(* IEC 61131-3 sources: plc-cip-batch-control/plc/types, 3 files *)

(* ---- Types_Cip.st ---- *)
(*
    Types_Cip.st: data types for the CIP skid controller.

    Naming follows the usual IEC prefixes: x BOOL, i INT, r REAL, t TIME,
    s STRING, e enumeration, st structure, fb function block instance.

    Enumeration members are prefixed because IEC 61131-3 puts them in the
    global namespace and PH_IDLE and UST_IDLE are different things.
*)

TYPE
    (* ISA-88 procedural state model, trimmed to the states this unit uses. *)
    E_UnitState : (
        UST_IDLE        := 0,
        UST_STARTING    := 1,
        UST_RUNNING     := 2,
        UST_HOLDING     := 3,
        UST_HELD        := 4,
        UST_RESTARTING  := 5,
        UST_COMPLETING  := 6,
        UST_COMPLETE    := 7,
        UST_ABORTING    := 8,
        UST_ABORTED     := 9
    );

    (* The CIP procedure. Phases run in this order; the recipe may skip some. *)
    E_Phase : (
        PH_IDLE                := 0,
        PH_PRE_RINSE           := 1,
        PH_CAUSTIC_WASH        := 2,
        PH_INTERMEDIATE_RINSE  := 3,
        PH_ACID_WASH           := 4,
        PH_FINAL_RINSE         := 5,
        PH_SANITISE            := 6,
        PH_COMPLETE            := 7
    );

    (* Every phase runs the same four steps; only its parameters differ. *)
    E_PhaseStep : (
        PS_IDLE      := 0,
        PS_LINEUP    := 1,
        PS_CHARGE    := 2,
        PS_CIRCULATE := 3,
        PS_RECOVER   := 4,
        PS_DONE      := 5
    );

    E_Source : (
        SRC_NONE       := 0,
        SRC_FRESH      := 1,
        SRC_RECOVERED  := 2,
        SRC_CAUSTIC    := 3,
        SRC_ACID       := 4
    );

    E_Return : (
        RET_DRAIN     := 0,
        RET_RECOVERY  := 1,
        RET_CAUSTIC   := 2,
        RET_ACID      := 3,
        RET_BALANCE   := 4
    );

    E_FailCode : (
        FC_NONE             := 0,
        FC_LINEUP_TIMEOUT   := 1,
        FC_CHARGE_TIMEOUT   := 2,
        FC_TEMP_TIMEOUT     := 3,
        FC_PHASE_TIMEOUT    := 4,
        FC_FLOW_LOW         := 5,
        FC_PUMP_FAULT       := 6,
        FC_OPERATOR_ABORT   := 7,
        FC_SAFETY_TRIP      := 8,
        FC_RINSE_NOT_CLEAN  := 9,
        FC_LEVEL_LOW        := 10,
        FC_SENSOR_FAULT     := 11
    );
END_TYPE

TYPE
    (*
        What one phase has to achieve. PRG_Sequence fills this from the recipe
        and hands it to the single phase engine, so adding a phase is a matter
        of parameters rather than another copy of the same logic.
    *)
    ST_PhaseParams : STRUCT
        eSource         : E_Source;
        eReturn         : E_Return;
        rTempSp         : REAL;     (* heat setpoint, degC *)
        rTempMin        : REAL;     (* below this the hold timer does not count *)
        rConcSp         : REAL;     (* chemical strength, % w/w *)
        rConcMin        : REAL;
        rConcMax        : REAL;
        rFlowSp         : REAL;     (* m3/h *)
        rFlowMin        : REAL;     (* below this the hold timer does not count *)
        tHold           : TIME;     (* verified hold required to pass *)
        tMinPhase       : TIME;
        tMaxPhase       : TIME;
        tRecover        : TIME;     (* push the circuit contents back or to drain *)
        xHeat           : BOOL;
        xDose           : BOOL;
        xRecirculate    : BOOL;     (* closed loop through the balance tank *)
        xAdaptiveEnd    : BOOL;     (* terminate on the return conductivity *)
        rEndConductivity : REAL;    (* mS/cm, adaptive rinses only *)
    END_STRUCT

    (* What the phase engine asks the control layer to do this scan. *)
    ST_Demand : STRUCT
        eSource      : E_Source;
        eReturn      : E_Return;
        rFlowSp      : REAL;
        rTempSp      : REAL;
        xHeat        : BOOL;
        xDose        : BOOL;
        xSupplyPump  : BOOL;
        xReturnPump  : BOOL;
        xFillValve   : BOOL;
    END_STRUCT

    (* One line of the electronic batch record. *)
    ST_PhaseResult : STRUCT
        ePhase           : E_Phase;
        xExecuted        : BOOL;
        xPass            : BOOL;
        eFail            : E_FailCode;
        rDurationS       : REAL;
        rHoldAchievedS   : REAL;
        rHoldRequiredS   : REAL;    (* zero when the endpoint is the conductivity *)
        xAdaptiveEnd     : BOOL;
        rMinTempC        : REAL := 999.0;
        rMaxTempC        : REAL;
        rMeanConcPct     : REAL;
        rMinFlow         : REAL := 999.0;
        rWaterL          : REAL;
        rChemL           : REAL;
        rEnergyKWh       : REAL;
        rEndConductivity : REAL;
    END_STRUCT

    ST_Recipe : STRUCT
        sName            : STRING[24] := 'default';
        xUseAcid         : BOOL := TRUE;
        xUseSanitise     : BOOL := FALSE;
        xAdaptive        : BOOL := FALSE;
        rFlowSp          : REAL := 18.0;
        tPreRinse        : TIME := T#3m;
        rCausticTempSp   : REAL := 75.0;
        rCausticTempMin  : REAL := 70.0;
        rCausticConcSp   : REAL := 2.0;
        tCausticHold     : TIME := T#10m;
        tIntRinse        : TIME := T#2m;
        rAcidTempSp      : REAL := 60.0;
        rAcidTempMin     : REAL := 55.0;
        rAcidConcSp      : REAL := 1.0;
        tAcidHold        : TIME := T#5m;
        tFinalRinse      : TIME := T#3m;
        rSanitiseTempSp  : REAL := 85.0;
        rSanitiseTempMin : REAL := 80.0;
        tSanitiseHold    : TIME := T#10m;
        rRinseEndCond    : REAL := 0.10;
        tPhaseMax        : TIME := T#45m;
        tRinseMax        : TIME := T#12m;   (* adaptive rinses fail rather than run on *)
        tRinseMin        : TIME := T#60s;   (* floor under the transport-delay blanking *)
        rFlowMin         : REAL := 14.0;
    END_STRUCT

    ST_Kpi : STRUCT
        rFreshWaterL     : REAL;
        rRecoveredWaterL : REAL;
        rEffluentL       : REAL;
        rCausticL        : REAL;
        rAcidL           : REAL;
        rEnergyKWh       : REAL;
        rCycleTimeS      : REAL;
        xVerifiedClean   : BOOL;
    END_STRUCT

    ST_Alarm : STRUCT
        xActive   : BOOL;
        xLatched  : BOOL;
        xAcked    : BOOL;
        iPriority : INT;
        rTimeInS  : REAL;
        iCount    : INT;
    END_STRUCT
END_TYPE

(* ---- GVL_Cip.st ---- *)
(*
    GVL_Cip.st: internal state shared between the five programs.

    Nothing here is located: these are the controller's own working data, not
    field I/O. PRG_Sequence owns the state and phase variables, PRG_Control owns
    the outputs, PRG_Alarms owns the alarm array and PRG_Kpi owns the totals.
    Every other program reads them.
*)

VAR_GLOBAL CONSTANT
    C_ALARM_COUNT       : INT  := 13;
    C_PHASE_COUNT       : INT  := 6;

    (* Alarm identifiers, used as the index into gAlarms. *)
    C_ALM_SAFETY        : INT  := 1;
    C_ALM_SUPPLY_PUMP   : INT  := 2;
    C_ALM_RETURN_PUMP   : INT  := 3;
    C_ALM_LEVEL_LOW     : INT  := 4;
    C_ALM_CAUSTIC_LOW   : INT  := 5;
    C_ALM_ACID_LOW      : INT  := 6;
    C_ALM_TEMP_LOW      : INT  := 7;
    C_ALM_FLOW_LOW      : INT  := 8;
    C_ALM_CIRCUIT_BUSY  : INT  := 9;
    C_ALM_PHASE_TIMEOUT : INT  := 10;
    C_ALM_NOT_CLEAN     : INT  := 11;
    C_ALM_NO_STEAM      : INT  := 12;
    C_ALM_COND_SENSOR   : INT  := 13;

    (* Skid geometry. The plant model holds the same figures; docs/model.md
       explains why they are stated twice and how the test keeps them equal. *)
    C_BALANCE_TANK_L    : REAL := 1200.0;
    C_CIRCUIT_VOLUME_L  : REAL := 450.0;    (* holdup of the circuit being cleaned *)
    (* A rinse endpoint cannot be believed until the return sensor has seen
       what was in the circuit when the rinse started. One and a half circuit
       turnovers is the blanking time. *)
    C_RINSE_TURNOVERS   : REAL := 1.5;
    C_FILL_TARGET_PCT   : REAL := 60.0;     (* recirculating phases *)
    (* Single-pass phases run the tank as a break volume at the lowest level
       the suction will stand. The rinse has to wash the tank out as well as
       the circuit and the tank washes out with a time constant of
       volume/flow: 156 litres at 18 m3/h is half a minute, 360 litres is
       nearly two and that difference is most of the rinse. *)
    C_RINSE_LEVEL_PCT   : REAL := 13.0;
    C_PUMP_START_PCT    : REAL := 10.0;     (* suction head to start the pump *)
    C_LEVEL_TRIP_PCT    : REAL := 7.0;
    C_CHEM_LEVEL_MIN    : REAL := 15.0;

    (* Two-point conductivity calibrations, mS/cm per % w/w, compensated to
       25 degC by the transmitter. Caustic is calibrated at 2 %, acid at 1 %. *)
    C_COND_K_CAUSTIC    : REAL := 47.0;
    C_COND_K_ACID       : REAL := 45.0;

    (* Positive-displacement dosing pumps, so the delivered volume is the
       valve-open time multiplied by a constant. *)
    C_CAUSTIC_DOSE_LPM  : REAL := 30.0;
    C_ACID_DOSE_LPM     : REAL := 20.0;

    C_TEMP_TOL          : REAL := 1.0;
    (* Plate-pack outlet limit. Above this the gaskets suffer and dissolved
       soil starts to bake onto the plates. *)
    C_SUPPLY_TEMP_LIMIT : REAL := 90.0;
    (* Task period. The harness asserts that the scan it runs matches. *)
    C_CYCLE_S           : REAL := 0.2;

    C_PUMP_SPEED_MIN    : REAL := 25.0;
    C_PUMP_SPEED_MAX    : REAL := 100.0;
END_VAR

VAR_GLOBAL
    (* ---- recipe and procedure state --------------------------------- *)
    gRecipe         : ST_Recipe;
    gUnitState      : E_UnitState;
    gPhase          : E_Phase;
    gPhaseStep      : E_PhaseStep;
    gFailCode       : E_FailCode;
    gPhaseParams    : ST_PhaseParams;
    gDemand         : ST_Demand;
    gResults        : ARRAY[1..6] OF ST_PhaseResult;
    gKpi            : ST_Kpi;
    giBatchId       : INT;

    (* ---- requests between programs ---------------------------------- *)
    gxSafetyTrip    : BOOL;     (* PRG_Safety -> everyone *)
    gxPermitRun     : BOOL;     (* PRG_Safety: it is safe to circulate *)
    gxPermitHeat    : BOOL;     (* PRG_Safety: steam may be admitted *)
    gxPermitDose    : BOOL;     (* PRG_Safety: chemical may be dosed *)
    gxHoldRequest   : BOOL;
    gxAbortRequest  : BOOL;
    gxPhaseExecute  : BOOL;
    gxPhaseDone     : BOOL;
    gxPhaseFailed   : BOOL;
    gxCycleReset    : BOOL;     (* one scan at the start of a batch *)
    gxPhaseStartPulse : BOOL;
    gxPhaseEndPulse : BOOL;
    giPhaseIndex    : INT;      (* which gResults entry the pulse refers to *)

    (* ---- derived measurements --------------------------------------- *)
    grConcentrationPct : REAL;  (* from the return conductivity *)
    grDeltaConductivity : REAL; (* return minus supply, the rinse criterion *)
    grCycleElapsedS : REAL;
    grPhaseElapsedS : REAL;
    grHoldAchievedS : REAL;
    grPlcTimeS      : REAL;     (* controller uptime, used to stamp alarms *)
    grCondFloor     : REAL;     (* reading the return must exceed in a wash *)
    gxCondSensorFault : BOOL;   (* the return element is not reading the process *)
    gxCondProven    : BOOL;     (* it saw the wash during this phase *)

    (* ---- alarms ------------------------------------------------------ *)
    gAlarms         : ARRAY[1..13] OF ST_Alarm;
    giFirstOut      : INT;
    giActiveAlarms  : INT;
    gxAlarmP1Active : BOOL;
END_VAR

(* ---- GVL_Io.st ---- *)
(*
    GVL_Io.st: the I/O image.

    These declarations are the single source of truth for the address map. The
    simulated field bus and the Modbus TCP server both build their tables by
    reading the AT addresses back out of the compiled program, so a tag cannot
    drift away from the address the logic uses. See docs/io_map.md.

    Address convention: %IXb.i is byte b bit i; %ID/%QD/%MD n is double word n.

    Inputs and outputs never share a number: inputs own bytes 0 and 1 and
    double words 0 to 15, outputs start at byte 2 and double word 16. IEC
    61131-3 keeps %I and %Q apart but some runtimes back both with one
    process image keyed by the number alone (RuSTy does, see
    docs/compiled_crosscheck.md); there %IX0.0 and %QX0.0 would be the same
    bit. Keeping the numbers disjoint costs nothing and works on both kinds.
*)

VAR_GLOBAL
    (* ---- digital inputs: plant status ------------------------------- *)
    xSafetyOk               AT %IX0.0 : BOOL;   (* safety relay healthy, E-stop clear *)
    xSupplyPumpRunning      AT %IX0.1 : BOOL;
    xReturnPumpRunning      AT %IX0.2 : BOOL;
    xSupplyPumpFault        AT %IX0.3 : BOOL;
    xReturnPumpFault        AT %IX0.4 : BOOL;
    xCircuitAvailable       AT %IX0.5 : BOOL;   (* the vessel is released for cleaning *)
    xSteamAvailable         AT %IX0.6 : BOOL;
    xBalanceTankLowLow      AT %IX0.7 : BOOL;   (* hard-wired float switch *)

    (* ---- operator commands -------------------------------------------
       These live in the memory area, not the input image, because they arrive
       from a panel or a SCADA client over the network rather than from a
       hard-wired button. The controller clears each one once it has taken the
       edge, so a client that writes a coil and forgets it still gets a pulse. *)
    xCmdStart               AT %MX0.0 : BOOL;
    xCmdHold                AT %MX0.1 : BOOL;
    xCmdRestart             AT %MX0.2 : BOOL;
    xCmdAbort               AT %MX0.3 : BOOL;
    xCmdReset               AT %MX0.4 : BOOL;
    xCmdAckAlarms           AT %MX0.5 : BOOL;

    (* ---- analogue inputs -------------------------------------------- *)
    rLevelBalanceTankPct    AT %ID0  : REAL;
    rTempSupplyC            AT %ID1  : REAL;    (* after the heat exchanger *)
    rTempReturnC            AT %ID2  : REAL;    (* back from the circuit *)
    rFlowSupplyM3h          AT %ID3  : REAL;
    rConductivityReturn     AT %ID4  : REAL;    (* mS/cm, temperature compensated *)
    rPressureSupplyBar      AT %ID5  : REAL;
    rLevelCausticPct        AT %ID6  : REAL;
    rLevelAcidPct           AT %ID7  : REAL;
    rLevelRecoveryPct       AT %ID8  : REAL;
    rConductivitySupply     AT %ID9  : REAL;    (* mS/cm, feed side *)
    rFlowMakeupM3h          AT %ID10 : REAL;    (* make-up into the balance tank *)
    rTempBalanceTankC       AT %ID11 : REAL;
    rConductivityTank       AT %ID12 : REAL;    (* CT-03, in the balance tank *)

    (* ---- digital outputs: valve matrix ------------------------------ *)
    xV01FreshWater          AT %QX2.0 : BOOL;
    xV02RecoveredWater      AT %QX2.1 : BOOL;
    xV03CausticDose         AT %QX2.2 : BOOL;
    xV04AcidDose            AT %QX2.3 : BOOL;
    xV05SupplyToCircuit     AT %QX2.4 : BOOL;
    xV06ReturnToDrain       AT %QX2.5 : BOOL;
    xV07ReturnToBalance     AT %QX2.6 : BOOL;
    xV08ReturnToCaustic     AT %QX2.7 : BOOL;
    xV09ReturnToRecovery    AT %QX3.0 : BOOL;
    xV10ReturnToAcid        AT %QX3.1 : BOOL;
    xSupplyPumpRun          AT %QX3.2 : BOOL;
    xReturnPumpRun          AT %QX3.3 : BOOL;
    xSteamIsolation         AT %QX3.4 : BOOL;
    xV11CausticSupply       AT %QX3.5 : BOOL;   (* caustic tank -> balance tank *)
    xV12AcidSupply          AT %QX3.6 : BOOL;

    (* ---- analogue outputs ------------------------------------------- *)
    rSupplyPumpSpeedPct     AT %QD16 : REAL;
    rSteamValvePct          AT %QD17 : REAL;

    (* ---- memory image published to SCADA ---------------------------- *)
    iHmiUnitState           AT %MW0 : INT;
    iHmiPhase               AT %MW1 : INT;
    iHmiPhaseStep           AT %MW2 : INT;
    iHmiFailCode            AT %MW3 : INT;
    iHmiActiveAlarms        AT %MW4 : INT;
    iHmiFirstOutAlarm       AT %MW5 : INT;
    iHmiBatchId             AT %MW6 : INT;

    rHmiFreshWaterL         AT %MD10 : REAL;
    rHmiRecoveredWaterL     AT %MD11 : REAL;
    rHmiEffluentL           AT %MD12 : REAL;
    rHmiCausticL            AT %MD13 : REAL;
    rHmiAcidL               AT %MD14 : REAL;
    rHmiEnergyKWh           AT %MD15 : REAL;
    rHmiCycleTimeS          AT %MD16 : REAL;
    rHmiPhaseElapsedS       AT %MD17 : REAL;
    rHmiHoldAchievedS       AT %MD18 : REAL;
    rHmiConcentrationPct    AT %MD19 : REAL;

    xHmiVerifiedClean       AT %MX30.0 : BOOL;
    xHmiCycleComplete       AT %MX30.1 : BOOL;
    xHmiCycleAborted        AT %MX30.2 : BOOL;
    xHmiAlarmHorn           AT %MX30.3 : BOOL;
    xHmiHeating             AT %MX30.4 : BOOL;
END_VAR
